(* CODESYS project BODAS-RC18-12_27-18_40-PR4.library
   Company: Bosch Rexroth AG
   DefaultNamespace: BODAS-RC18-12_27-18_40-PR4
   Title: BODAS_RC18-12_27-18_40-PR4
   DocFormat: reStructuredText
   Description: User library to use BODAS-BDL services (API) for RC40.
   Version: 2.3.0

Project tree, tasks and I/O mapping:
  PR4/
    API/
      function bds_snsrPr4_getPressure [ST]
      function bds_snsrPr4_getTemp [ST]
    ENUM/
      data type bds_snsrPr4_status_te
    UNION/
      data type bds_snsrPr4_statusDiag_tu
    STRUCT/
      data type bds_snsrPr4_getPressure_ts
      data type bds_snsrPr4sent_statusDiag_tb
      data type bds_snsrPr4_getTemp_ts
      data type bds_snsrPr4an_statusDiag_tb
*)

// PR4/ENUM/bds_snsrPr4_status_te
{attribute 'external_name' := 'cmp_rts_bds_snsrPr4_status_te'}
TYPE bds_snsrPr4_status_te :
(
	bds_snsrPr4_ok_E := 0,
	bds_snsrPr4_init_E := 1,
	bds_snsrPr4_noUpdate_E := 2,
	bds_snsrPr4_outOfRange_E := 3,
	bds_snsrPr4_err_E := 4,
	bds_snsrPr4_invldConfig_E := 5,
	bds_snsrPr4_invldPrm_E := 6
)USINT;
END_TYPE

// PR4/STRUCT/bds_snsrPr4_getPressure_ts
{attribute 'external_name' := 'cmp_rts_bds_snsrPr4_getPressure_ts'}
TYPE bds_snsrPr4_getPressure_ts :
STRUCT
	stsApi_e: bds_snsrPr4_status_te;  // stsApi_e			   Status of the BDL API function call.
	pressureMeasmtRng_dBar_u16: UINT; // Return of the pressure measurement range value from 0 deci bar to the determined value of the Pr4 sensor with resolution in deci bar
	statusDiag_u: bds_snsrPr4_statusDiag_tu; // statusDiag_u 	       Status diagnostic information of Pr4 sensor.
	pressure_dBar_u16: UINT; //	pressure_dBar_u16	   Measured pressure value FROM Pr4 sensor with resolution in deci bar.
	padding: ARRAY[0..1] OF BYTE;  // Add 2 bytes padding
END_STRUCT
END_TYPE

// PR4/STRUCT/bds_snsrPr4sent_statusDiag_tb
(*Bit field type definition for the output module with diagnostic status information of output pin.*)
{attribute 'external_name' := 'cmp_rts_bds_snsrPr4sent_statusDiag_tb'}
{attribute 'size' := '32'}
 
TYPE bds_snsrPr4sent_statusDiag_tb :
STRUCT
	stErrSnsr_b1: BIT; /// stErrSCB_b1 Fault error status bit information for;·pressure or temperature above or below limit or overflows or saturation in supply voltage path (measurement possibly unreliable or wrong) or overflows or saturation in signal paths (pressure, temperature, supply voltage).
	stErrVdd_b1: BIT; // stErrVdd_b1 :  Fault error status bit information for low or high thresholds voltage supply exceeded.
	resd1_b : ARRAY[0..2] OF BYTE;      (* Reserved *)
END_STRUCT
END_TYPE

// PR4/STRUCT/bds_snsrPr4_getTemp_ts
{attribute 'external_name' := 'cmp_rts_bds_snsrPr4_getTemp_ts'}
TYPE bds_snsrPr4_getTemp_ts :
STRUCT
	stsApi_e: bds_snsrPr4_status_te;  // tatus of the BDL API function call
	statusDiag_u: bds_snsrPr4_statusDiag_tu; // Status diagnostic information of Pr4 sensor.
	temp_degC_s32: DINT; // Measured pressure value from Pr4 sensor with resolution in deci bar.
END_STRUCT
END_TYPE

// PR4/STRUCT/bds_snsrPr4an_statusDiag_tb
(*Bit field type definition for the output module with diagnostic status information of output pin.*)
{attribute 'external_name' := 'cmp_rts_bds_snsrPr4an_statusDiag_tb'}
{attribute 'size' := '32'}

TYPE bds_snsrPr4an_statusDiag_tb :
STRUCT
	stErrSCB_b1: BIT;   // stErrSCB_b1 Fault error status for short cut to battery
	stErrSCG_b1: BIT;   // stErrSCG_b1 :  Fault error status for short cut to ground
	stErrOL_b1: BIT;    // stErrOL_b1 : Fault error status for open load
	stErrHw_b1: BIT;    // stErrHw_b1 : Fault error status for hardware error for example  ADC connection is broken.
	resd1_b : ARRAY[0..2] OF BYTE;      (* Reserved *)
END_STRUCT
END_TYPE

// PR4/UNION/bds_snsrPr4_statusDiag_tu
{attribute 'external_name' := 'cmp_rts_bds_snsrPr4_statusDiag_tu'}
TYPE bds_snsrPr4_statusDiag_tu :

UNION
	anStDiag_b: bds_snsrPr4an_statusDiag_tb;
	sentStDiag_b: bds_snsrPr4sent_statusDiag_tb;
END_UNION

END_TYPE

// PR4/API/bds_snsrPr4_getPressure
/// The bds_snsrPr4_getPressure API function provides calculated pressure with resolution of deci bar and diagnostic status of a particular PR4 sensor instance.
///
///Remarks
///
///A configuration of the PR4 SENT sensor type is necessary and this will be done automatically with the received SENT slow data message with the message ID 0x08 from the PR4 SENT sensor.
///
///  
///==================================================================		  			===================================================================================================
///Return value    								  									     Description
///==================================================================		  			===================================================================================================
/// bds_snsrPr4_getPressure_ts															The return structure containing the status of API function call, pressure in deci-bar and diagnostic information of a particular PR4 sensor instance. For detail information please refer into chapter PR4 SENT.																
///
///==================================================================		   			===================================================================================================
///
///=======
///Code Example:
///=======
///============================================================================
///
/// PROGRAM appl_10ms_task
/// 
/// VAR
/// 
///     bds_snsrPr4_getPressure_s: bds_snsrPr4_getPressure_ts;
/// 	
///     bds_snsrPr4_inst_e: bds_snsrPr4_inst_te;
/// 	
///     pressureLocal_dBar_u16: UINT;  (* pressure in deci-bar *)
/// 	
/// END_VAR
/// 
/// (* PR4 sensor instance *)
/// 
/// bds_snsrPr4_inst_e := bds_snsrPr4_inst_te.PumpPressure_E;
/// 
/// (* BDL API function call *)
/// 
/// bds_snsrPr4_getPressure_s := bds_snsrPr4_getPressure(bds_snsrPr4_inst_e);
/// 
/// (* check the return status of API function call *)
/// 
/// IF bds_snsrPr4_ok_E = bds_snsrPr4_getPressure_s.stsApi_e THEN
/// 
///     (* save the actual wheel speed and rotation direction *)
/// 	
///     pressureLocal_dBar_u16 := bds_snsrPr4_getPressure_s.pressure_dBar_u16;
/// 	
/// ELSE
/// 
///     (* error handling *)
/// 	
/// END_IF
/// 
/// END_PROGRAM
///
///============================================================================
{attribute 'external_name' := 'cmp_rts_bds_snsrPr4_getPressure'}
FUNCTION bds_snsrPr4_getPressure : bds_snsrPr4_getPressure_ts
VAR_INPUT
	/// The PR4 sensor instance name.
	snsrPr4Inst_e: USINT;
END_VAR

END_FUNCTION

// PR4/API/bds_snsrPr4_getTemp
/// The bds_snsrPr4_getPressure API function provides calculated pressure with resolution of deci bar and diagnostic status of a particular PR4 sensor instance.
///
///Remarks
///
///A configuration of the PR4 SENT sensor type is necessary and this will be done automatically with the received SENT slow data message with the message ID 0x08 from the PR4 SENT sensor.
///
///  
///==================================================================		  			===================================================================================================
///Return value    								  									     Description
///==================================================================		  			===================================================================================================
/// bds_snsrPr4_getTemp_ts															    The return structure containing the status of API function call, temperature in degree Celsius and diagnostic information of a particular PR4 sensor instance. For detail information please refer into chapter PR4 SENT.																
///
///==================================================================		   			===================================================================================================
///
///=======
///Code Example:
///=======
///============================================================================
///
/// PROGRAM appl_10ms_task
/// 
/// VAR
/// 
///     bds_snsrPr4_getTemp_s : bds_snsrPr4_getTemp_ts;
/// 	
///     bds_snsrPr4_inst_e : bds_snsrPr4_inst_te;
/// 	
///     temp_degC_s32 : DINT;  
/// 	
/// END_VAR
/// 
/// (* PR4 sensor instance *)
/// 
/// bds_snsrPr4_inst_e := bds_snsrPr4_inst_te.PumpPressure_E;
/// 
/// (* BDL API function call *)
/// 
/// bds_snsrPr4_getTemp_s := bds_snsrPr4_getTemp(bds_snsrPr4_inst_e);
/// 
/// (* Check the return status of API function call *)
/// 
/// IF bds_snsrPr4_getTemp_s.stsApi_e = bds_snsrPr4_ok_E THEN
/// 
///     (* Save the actual temperature in degree celsius *)
/// 	
///     temp_degC_s32 := bds_snsrPr4_getTemp_s.temp_degC_s32;
/// 	
/// ELSE
/// 
///     (* Error handling *)
/// 	
///     (* Add your error handling code here *)
/// 	
/// END_IF;

/// END_PROGRAM
///
///============================================================================
{attribute 'external_name' := 'cmp_rts_bds_snsrPr4_getTemp'}
FUNCTION bds_snsrPr4_getTemp : bds_snsrPr4_getTemp_ts
VAR_INPUT
	/// The PR4 sensor instance name.
	snsrPr4Inst_e: USINT;
END_VAR

END_FUNCTION
